// Mitsubishi GX Works2 project: 260928_기초회로_잠등지연   PLC: Q03UDV

PROGRAM MAIN
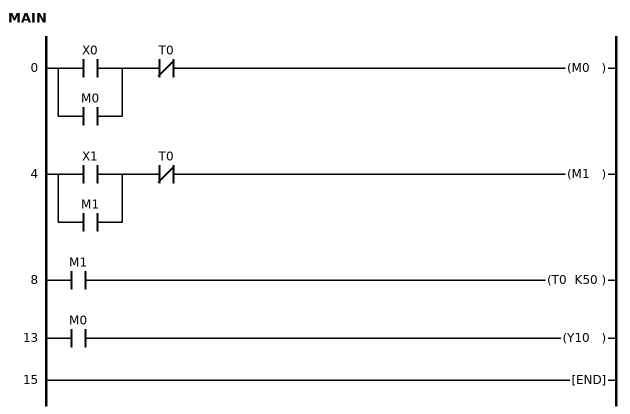
0     LD      X0
      OR      M0
      ANI     T0
      OUT     M0
4     LD      X1
      OR      M1
      ANI     T0
      OUT     M1
8     LD      M1
      OUT     T0 K50
13    LD      M0
      OUT     Y10
15    END
END_PROGRAM
